(* PLC project probe, plc-portfolio cds2astra probe 0.1.0 *)
(* stored: creationDateTime 2026-10-20T00:00:00, modificationDateTime 2026-10-20T00:00:00 *)

PROGRAM PRG_P4
VAR
    xA : BOOL;
    xQ : BOOL;
END_VAR

            LD xA
NOT
ST xQ

          
END_PROGRAM
